(* Logix 5000 project; controller SEAS_475 vendor 1 type 14 code 77 rev 17.4; software revision 17.01 *)

TASK MainTask (continuous, watchdog 500 ms) : MainProgram

MODULES
   Controller : vendor 1 type 14 code 77 (CompactLogixL32EController 0, rev 17.4)
      LocalENB : 1769-L32E Ethernet Port (CompactLogixL32Ethernet 1, rev 17.2)
         robot : ETHERNET-MODULE (Ethernet 192.168.1.100, rev 1.1, Output RPI 10 ms)
      Local : CompactBus (CompactVirtualAdapter 3, rev 17.2, Input RPI 5 ms)
         Input_Output1 : vendor 1 type 7 code 66 (Compact 4, rev 2.1, Output RPI 5 ms)
         Input_Output2 : vendor 1 type 7 code 66 (Compact 5, rev 2.1, Output RPI 5 ms)
         Input_1 : 1769-IQ16 (Compact 1, rev 1.1, Input RPI 5 ms)
         Input_2 : 1769-IQ16 (Compact 2, rev 1.1, Input RPI 5 ms)
         Output_1 : 1769-OB16 (Compact 3, rev 2.1, Output RPI 5 ms)
         Output_2 : 1769-OB16 (Compact 6, rev 2.1, Output RPI 5 ms)
END_MODULES

VAR_GLOBAL   (* controller tags *)
   b1 : DINT;
   B2 : DINT;
   B3_10_Fanuc_Produced_DIN_3 : DINT; {produced}
   B3_11_Fanuc_Produced_DOUT_3 : DINT; {produced}
   B3_12_Fanuc_Produced_DIN_4 : DINT; {produced}
   B3_13_Fanuc_Produced_DOUT_4 : DINT; {produced}
   B3_2_L32_Produced_Outputs_1 : DINT := 327682; {produced}
   B3_3_L32_Produced_Inputs_1 : DINT := 131074; {produced}
   B3_4_L32_Produced_Output_2 : DINT; {produced}
   B3_5_L32_Produced_Inputs_2 : DINT; {produced}
   B3_6_Fanuc_Produced_DIN_1 : DINT := 135; {produced}
   B3_7_Fanuc_Produced_DOUT_1 : DINT := 160; {produced}
   B3_8_Fanuc_Produced_DIN_2 : DINT; {produced}
   B3_9_Fanuc_Produced_DOUT_2 : DINT; {produced}
   C1 : COUNTER := (PRE := 1, ACC := 5, CU := 1, DN := 1);
   C2 : COUNTER := (PRE := 4, ACC := 21, DN := 1);
   Data_Start : DINT; {produced}
   Db_Stop : DINT; {produced}
   IMU_Tare : DINT; {produced}
   Pause_Bit : DINT;
   push_button_1_timer : TIMER := (PRE := 10000, ACC := 10000, EN := 1, DN := 1);
   PUSH_BUTTON_BITS : DINT;
   t1 : TIMER := (PRE := 300);
   t2 : TIMER := (PRE := 100);
   t3 : TIMER := (PRE := 200);
   t4 : TIMER := (PRE := 300);
END_VAR

PROGRAM MainProgram   (* main routine MainRoutine *)
VAR
   Fanuc_Invis : BOOL;
   Fanuc_Mov : COUNTER := (PRE := 1, ACC := 1, DN := 1);
   Fanuc_Mov_Cam1 : TIMER := (PRE := 40000, ACC := 40000, EN := 1, DN := 1);
   Fanuc_Mov_Perch : TIMER := (PRE := 27000, ACC := 27000, EN := 1, DN := 1);
   Fanuc_mov_Steve : TIMER := (PRE := 40000);
   Fanuc_Rot_invs : BOOL := 1;
   Fanuc_Stationary : BOOL;
   HMI_Reset_Light : BOOL := 1;
   Reset_for_HMI : BOOL;
   Start_for_HMI : BOOL;
   steve_arm1_invis : BOOL := 1;
   steve_arm2_invis : BOOL := 1;
   steve_mov_bk : TIMER := (PRE := 25000, ACC := 25000, EN := 1, DN := 1);
   Steve_Move_Timer : TIMER := (PRE := 15000, ACC := 15000, EN := 1, DN := 1);
   Steve_perch : BOOL;
   Stop_for_HMI : BOOL;
   System_Ready_HMI : BOOL;
END_VAR

ROUTINE MainRoutine   (* ladder *)
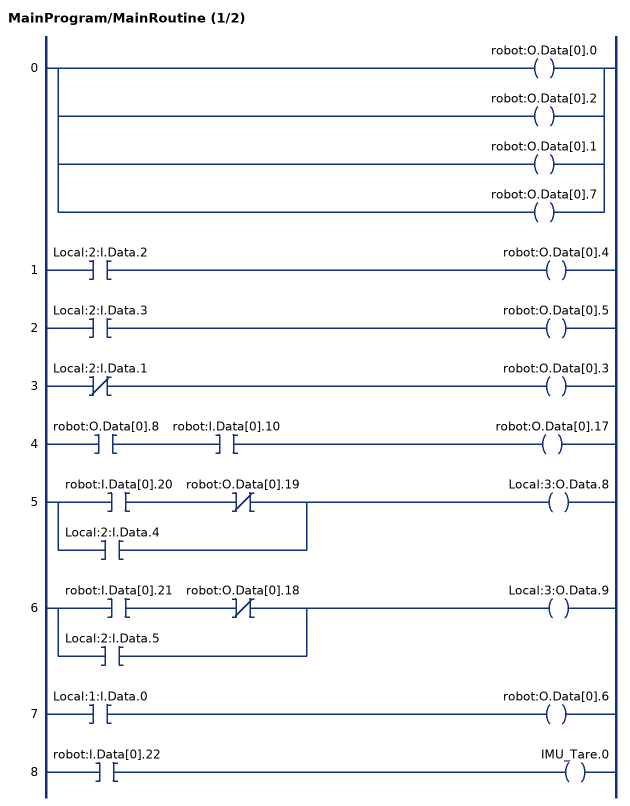
   0: [OTE(robot:O.Data[0].0) ,[OTE(robot:O.Data[0].2) ,[OTE(robot:O.Data[0].1) ,OTE(robot:O.Data[0].7) ] ] ];
   1: XIC(Local:2:I.Data.2)OTE(robot:O.Data[0].4);
   2: XIC(Local:2:I.Data.3)OTE(robot:O.Data[0].5);
   3: XIO(Local:2:I.Data.1)OTE(robot:O.Data[0].3);
   4: XIC(robot:O.Data[0].8)XIC(robot:I.Data[0].10)OTE(robot:O.Data[0].17);
   5: [XIC(robot:I.Data[0].20) XIO(robot:O.Data[0].19) ,XIC(Local:2:I.Data.4) ]OTE(Local:3:O.Data.8);
   6: [XIC(robot:I.Data[0].21) XIO(robot:O.Data[0].18) ,XIC(Local:2:I.Data.5) ]OTE(Local:3:O.Data.9);
   7: XIC(Local:1:I.Data.0)OTE(robot:O.Data[0].6);
   8: XIC(robot:I.Data[0].22)OTE(IMU_Tare.0);
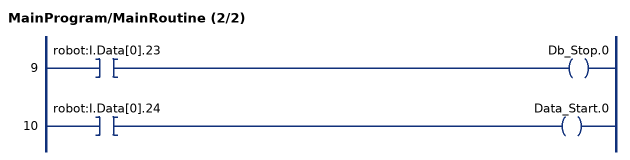
   9: XIC(robot:I.Data[0].23)OTE(Db_Stop.0);
   10: XIC(robot:I.Data[0].24)OTE(Data_Start.0);
END_ROUTINE
END_PROGRAM
